(* IEC 61131-3 sources: 2026_Projet_YGO_ExcavatriceDragage/TOOLS/TEST_AUTO_CI/RESULTS/H_TREUILS_BENNE/reports (part 5) *)

    machine(HeartbeatIhmOk := TRUE, CanBusOperational := TRUE, JoyOperational := TRUE, CmdMode := E_Mode.DISABLE, TglJoystickMaster := TRUE, JoyRawY := 8000, CmdWinchSelect := 1);
    ADVANCE_TIME(20000000);
    machine(HeartbeatIhmOk := TRUE, CanBusOperational := TRUE, JoyOperational := TRUE, TglJoystickMaster := TRUE, JoyRawY := 8000, CmdWinchSelect := 1);
    ASSERT_TRUE(machine.BusOutputs.M1RelayFwd = FALSE, 'HARN-71: Enable=FALSE -> sorties sures');
    ASSERT_EQ(machine.M1_StepNumber, 0, 'HARN-71: palier neutralise');

    machine(HeartbeatIhmOk := TRUE, CanBusOperational := TRUE, JoyOperational := TRUE, CmdMode := E_Mode.MAINT_N1, TglJoystickMaster := TRUE, JoyRawY := 8000, CmdWinchSelect := 1);
    ADVANCE_TIME(50000000);
    machine(HeartbeatIhmOk := TRUE, CanBusOperational := TRUE, JoyOperational := TRUE, TglJoystickMaster := TRUE, JoyRawY := 8000, CmdWinchSelect := 1);
    (* ORACLE (main) : la reprise exige une NOUVELLE intention — l'adoption immédiate
       au ré-Enable = défaut D18 (rouge baseline attendu, cible T181-05) *)
    ASSERT_TRUE(machine.BusOutputs.M1RelayFwd = FALSE, 'HARN-71: pas de redemarrage auto au re-Enable (cible D18)');
END_TEST

TEST 'HARN-72 : Watchdog frein (retour frein ne suit pas) -> barriere coupe apres timeout'
    seqReqM1.RunRequest := FALSE; seqReqM1.ReqAscent := FALSE; seqReqM1.StepTgt := 0;
    seqReqM2.RunRequest := FALSE; seqReqM2.ReqAscent := FALSE; seqReqM2.StepTgt := 0;
    seqReqBucket.ExtractionControlActive := FALSE; seqReqBucket.DescendPermitDiveBucketOpen := FALSE;
    machine(HeartbeatIhmOk := TRUE, CanBusOperational := TRUE, JoyOperational := TRUE,
        CmdMode := E_Mode.MAINT_N1, CmdWinchSelect := 1, TglJoystickMaster := TRUE,
        SpeedTable := speedTable, ModelStepSpeedMps := modelSpeeds,
        SeqReqWinchM1 := seqReqM1, SeqReqWinchM2 := seqReqM2, SeqReqBucket := seqReqBucket,
        ModelSeedPosM1 := 2.0, ModelSeedPosM2 := 2.0, ModelReloadPositions := TRUE,
        ModelM2SpeedFactor := 1.0,
        ModelBrakeFeedbackFaultM1 := TRUE, (* retour frein M1 ne s ouvre jamais *)
        JoyRawX := 5000, JoyRawY := 5000, JoyDeadmanBtn := FALSE,
        EmergencyChainClosed := TRUE, PowerContactorEngaged := TRUE, HeartbeatIhmOk := TRUE
    );
    (* T181-00b : retour neutre sans commande >= 1500 ms pour purger RestartRequired/DeadTime *)
    machine(HeartbeatIhmOk := TRUE, CanBusOperational := TRUE, JoyOperational := TRUE, JoyDeadmanBtn := TRUE, TglJoystickMaster := TRUE, JoyRawY := 5000, CmdWinchSelect := 1, CmdMode := E_Mode.MAINT_N1);
    ADVANCE_TIME(2000000000);
    machine(HeartbeatIhmOk := TRUE, CanBusOperational := TRUE, JoyOperational := TRUE, JoyDeadmanBtn := TRUE, TglJoystickMaster := TRUE, JoyRawY := 5000, CmdWinchSelect := 1, CmdMode := E_Mode.MAINT_N1);
    machine(HeartbeatIhmOk := TRUE, CanBusOperational := TRUE, JoyOperational := TRUE, JoyDeadmanBtn := TRUE, TglJoystickMaster := TRUE, JoyRawY := 8000, CmdWinchSelect := 1, CmdMode := E_Mode.MAINT_N1);
    ADVANCE_TIME(5000000000); (* 5 s : tout timeout frein realiste a expire *)
    machine(HeartbeatIhmOk := TRUE, CanBusOperational := TRUE, JoyOperational := TRUE, TglJoystickMaster := TRUE, JoyRawY := 8000, CmdWinchSelect := 1, CmdMode := E_Mode.MAINT_N1);

    (* ORACLE (main) : frein incohérent -> la barrière coupe la commande de sens (TC-P10-012) *)
    ASSERT_TRUE(machine.BusWinch.WinchM1FinalInterlockRequest.RequestedRelayFwd, 'HARN-72: FB_Winch demande toujours le sens (defaut cote barriere)');
    ASSERT_TRUE(machine.BusOutputs.M1RelayFwd = FALSE, 'HARN-72: barriere a coupe (watchdog frein)');
    ASSERT_TRUE(machine.FinalInterlockGovernedM1, 'HARN-72: FinalInterlockGoverned TRUE');
END_TEST

TEST 'HARN-73 : Temps mort directionnel apres arret (inversion 200 ms) -> RelayRev retenu (CIBLE T175/T181-05)'
    seqReqM1.RunRequest := FALSE; seqReqM1.ReqAscent := FALSE; seqReqM1.StepTgt := 0;
    seqReqM2.RunRequest := FALSE; seqReqM2.ReqAscent := FALSE; seqReqM2.StepTgt := 0;
    seqReqBucket.ExtractionControlActive := FALSE; seqReqBucket.DescendPermitDiveBucketOpen := FALSE;
    machine(HeartbeatIhmOk := TRUE, CanBusOperational := TRUE, JoyOperational := TRUE,
        CmdMode := E_Mode.MAINT_N1, CmdWinchSelect := 1, TglJoystickMaster := TRUE,
        SpeedTable := speedTable, ModelStepSpeedMps := modelSpeeds,
        SeqReqWinchM1 := seqReqM1, SeqReqWinchM2 := seqReqM2, SeqReqBucket := seqReqBucket,
        ModelSeedPosM1 := 2.0, ModelSeedPosM2 := 2.0, ModelReloadPositions := TRUE,
        ModelM2SpeedFactor := 1.0,
        JoyRawX := 5000, JoyRawY := 5000, JoyDeadmanBtn := FALSE,
        EmergencyChainClosed := TRUE, PowerContactorEngaged := TRUE, HeartbeatIhmOk := TRUE
    );
    (* T181-00b : retour neutre sans commande >= 1500 ms pour purger RestartRequired/DeadTime *)
    machine(HeartbeatIhmOk := TRUE, CanBusOperational := TRUE, JoyOperational := TRUE, JoyDeadmanBtn := TRUE, TglJoystickMaster := TRUE, JoyRawY := 5000, CmdWinchSelect := 1, CmdMode := E_Mode.MAINT_N1);
    ADVANCE_TIME(2000000000);
    machine(HeartbeatIhmOk := TRUE, CanBusOperational := TRUE, JoyOperational := TRUE, JoyDeadmanBtn := TRUE, TglJoystickMaster := TRUE, JoyRawY := 5000, CmdWinchSelect := 1, CmdMode := E_Mode.MAINT_N1);
    machine(HeartbeatIhmOk := TRUE, CanBusOperational := TRUE, JoyOperational := TRUE, JoyDeadmanBtn := TRUE, TglJoystickMaster := TRUE, JoyRawY := 8000, CmdWinchSelect := 1, CmdMode := E_Mode.MAINT_N1);
    ADVANCE_TIME(200000000);
    machine(HeartbeatIhmOk := TRUE, CanBusOperational := TRUE, JoyOperational := TRUE, TglJoystickMaster := TRUE, JoyRawY := 8000, CmdWinchSelect := 1, CmdMode := E_Mode.MAINT_N1);
    machine(HeartbeatIhmOk := TRUE, CanBusOperational := TRUE, JoyOperational := TRUE, JoyDeadmanBtn := TRUE, TglJoystickMaster := TRUE, JoyRawY := 5000, CmdWinchSelect := 1, CmdMode := E_Mode.MAINT_N1);
    ADVANCE_TIME(20000000);
    machine(HeartbeatIhmOk := TRUE, CanBusOperational := TRUE, JoyOperational := TRUE, TglJoystickMaster := TRUE, JoyRawY := 5000, CmdWinchSelect := 1, CmdMode := E_Mode.MAINT_N1);
    (* Inversion 200 ms après l'arrêt *)
    machine(HeartbeatIhmOk := TRUE, CanBusOperational := TRUE, JoyOperational := TRUE, JoyDeadmanBtn := TRUE, TglJoystickMaster := TRUE, JoyRawY := 2000, CmdWinchSelect := 1, CmdMode := E_Mode.MAINT_N1);
    ADVANCE_TIME(200000000);
    machine(HeartbeatIhmOk := TRUE, CanBusOperational := TRUE, JoyOperational := TRUE, TglJoystickMaster := TRUE, JoyRawY := 2000, CmdWinchSelect := 1, CmdMode := E_Mode.MAINT_N1);

    (* PRECOND (durcissement T181-00b) : la barriere ne doit etre testee que si la demande de
       descente est REELlement presente en amont (RequestedRelayRev). Sans elle, M1RelayRev=FALSE
       est une tautologie (aucune demande a retenir). *)
    ASSERT_TRUE(machine.BusWinch.WinchM1FinalInterlockRequest.RequestedRelayRev, 'HARN-73: precondition - inversion descente reellement demandee');
    (* ORACLE (main) : délai interlock descente (400 ms) non écoulé -> la barriere retient RelayRev *)
    ASSERT_TRUE(machine.BusOutputs.M1RelayRev = FALSE, 'HARN-73: temps mort directionnel respecte (cible T175)');
END_TEST

TEST 'HARN-74a : Coast-down apres relache lourd -> PAS de faux PowerCutOff pendant la fenetre contacteurs (T178)'
    seqReqM1.RunRequest := FALSE; seqReqM1.ReqAscent := FALSE; seqReqM1.StepTgt := 0;
    seqReqM2.RunRequest := FALSE; seqReqM2.ReqAscent := FALSE; seqReqM2.StepTgt := 0;
    seqReqBucket.ExtractionControlActive := FALSE; seqReqBucket.DescendPermitDiveBucketOpen := FALSE;
    machine(HeartbeatIhmOk := TRUE, CanBusOperational := TRUE, JoyOperational := TRUE,
        CmdMode := E_Mode.MAINT_N1, CmdWinchSelect := 1, TglJoystickMaster := TRUE,
        SpeedTable := speedTable, ModelStepSpeedMps := modelSpeeds,
        SeqReqWinchM1 := seqReqM1, SeqReqWinchM2 := seqReqM2, SeqReqBucket := seqReqBucket,
        ModelSeedPosM1 := 2.0, ModelSeedPosM2 := 2.0, ModelReloadPositions := TRUE,
        ModelM2SpeedFactor := 1.0,
        JoyRawX := 5000, JoyRawY := 8000, JoyDeadmanBtn := FALSE,
        EmergencyChainClosed := TRUE, PowerContactorEngaged := TRUE, HeartbeatIhmOk := TRUE
    );
    (* T181-00b : retour neutre sans commande >= 1500 ms pour purger RestartRequired/DeadTime *)
    machine(HeartbeatIhmOk := TRUE, CanBusOperational := TRUE, JoyOperational := TRUE, JoyDeadmanBtn := TRUE, TglJoystickMaster := TRUE, JoyRawY := 5000, CmdWinchSelect := 1, CmdMode := E_Mode.MAINT_N1);
    ADVANCE_TIME(2000000000);
    machine(HeartbeatIhmOk := TRUE, CanBusOperational := TRUE, JoyOperational := TRUE, JoyDeadmanBtn := TRUE, TglJoystickMaster := TRUE, JoyRawY := 5000, CmdWinchSelect := 1, CmdMode := E_Mode.MAINT_N1);
    machine(HeartbeatIhmOk := TRUE, CanBusOperational := TRUE, JoyOperational := TRUE, JoyDeadmanBtn := TRUE, TglJoystickMaster := TRUE, JoyRawY := 8000, CmdWinchSelect := 1, CmdMode := E_Mode.MAINT_N1);
    ADVANCE_TIME(200000000);
    machine(HeartbeatIhmOk := TRUE, CanBusOperational := TRUE, JoyOperational := TRUE, TglJoystickMaster := TRUE, JoyRawY := 8000, CmdWinchSelect := 1, CmdMode := E_Mode.MAINT_N1);
    ASSERT_TRUE(machine.BusOutputs.M1RelayFwd, 'HARN-74a: precondition - montee plein pot');

    (* Relâche homme-mort plein déflexion : coast 500 ms (contacteurs pas encore retombés, v > 0) *)
    machine(HeartbeatIhmOk := TRUE, CanBusOperational := TRUE, JoyOperational := TRUE, JoyDeadmanBtn := FALSE, TglJoystickMaster := TRUE, JoyRawY := 8000, CmdWinchSelect := 1, CmdMode := E_Mode.MAINT_N1);
    ADVANCE_TIME(100000000); (* 100 ms au coeur de la fenêtre coast *)
    machine(HeartbeatIhmOk := TRUE, CanBusOperational := TRUE, JoyOperational := TRUE, TglJoystickMaster := TRUE, JoyRawY := 8000, CmdWinchSelect := 1, CmdMode := E_Mode.MAINT_N1);

    (* ORACLE (main) : pendant le coast — mouvement résiduel SANS commande : Méca A ne doit PAS armer *)
    ASSERT_TRUE(machine.BusWinch.WinchM1Safety.PowerCutOff = FALSE, 'HARN-74a: PAS de faux PowerCutOff pendant le coast (T178)');
    ASSERT_TRUE(machine.BusWinch.WinchM1Safety.SafeStop = FALSE, 'HARN-74a: PAS de SafeStop pendant le coast (Meca A)');
END_TEST

TEST 'HARN-74b : Coast-down prolonge -> Meca B arme a 3 s (CIBLE T178, ROUGE baseline)'
    seqReqM1.RunRequest := FALSE; seqReqM1.ReqAscent := FALSE; seqReqM1.StepTgt := 0;
    seqReqM2.RunRequest := FALSE; seqReqM2.ReqAscent := FALSE; seqReqM2.StepTgt := 0;
    seqReqBucket.ExtractionControlActive := FALSE; seqReqBucket.DescendPermitDiveBucketOpen := FALSE;
    machine(HeartbeatIhmOk := TRUE, CanBusOperational := TRUE, JoyOperational := TRUE,
        CmdMode := E_Mode.MAINT_N1, CmdWinchSelect := 1, TglJoystickMaster := TRUE,
        SpeedTable := speedTable, ModelStepSpeedMps := modelSpeeds,
        SeqReqWinchM1 := seqReqM1, SeqReqWinchM2 := seqReqM2, SeqReqBucket := seqReqBucket,
        ModelSeedPosM1 := 2.0, ModelSeedPosM2 := 2.0, ModelReloadPositions := TRUE,
        ModelM2SpeedFactor := 1.0,
        JoyRawX := 5000, JoyRawY := 8000, JoyDeadmanBtn := FALSE,
        EmergencyChainClosed := TRUE, PowerContactorEngaged := TRUE, HeartbeatIhmOk := TRUE
    );
    (* T181-00b : retour neutre sans commande >= 1500 ms pour purger RestartRequired/DeadTime *)
    machine(HeartbeatIhmOk := TRUE, CanBusOperational := TRUE, JoyOperational := TRUE, JoyDeadmanBtn := TRUE, TglJoystickMaster := TRUE, JoyRawY := 5000, CmdWinchSelect := 1, CmdMode := E_Mode.MAINT_N1);
    ADVANCE_TIME(2000000000);
    machine(HeartbeatIhmOk := TRUE, CanBusOperational := TRUE, JoyOperational := TRUE, JoyDeadmanBtn := TRUE, TglJoystickMaster := TRUE, JoyRawY := 5000, CmdWinchSelect := 1, CmdMode := E_Mode.MAINT_N1);
    machine(HeartbeatIhmOk := TRUE, CanBusOperational := TRUE, JoyOperational := TRUE, JoyDeadmanBtn := TRUE, TglJoystickMaster := TRUE, JoyRawY := 8000, CmdWinchSelect := 1, CmdMode := E_Mode.MAINT_N1);
    ADVANCE_TIME(200000000);
    machine(HeartbeatIhmOk := TRUE, CanBusOperational := TRUE, JoyOperational := TRUE, TglJoystickMaster := TRUE, JoyRawY := 8000, CmdWinchSelect := 1, CmdMode := E_Mode.MAINT_N1);
    machine(HeartbeatIhmOk := TRUE, CanBusOperational := TRUE, JoyOperational := TRUE, JoyDeadmanBtn := FALSE, TglJoystickMaster := TRUE, JoyRawY := 8000, CmdWinchSelect := 1, CmdMode := E_Mode.MAINT_N1);
    ADVANCE_TIME(4000000000); (* 4 s > 3 s *)
    machine(HeartbeatIhmOk := TRUE, CanBusOperational := TRUE, JoyOperational := TRUE, TglJoystickMaster := TRUE, JoyRawY := 8000, CmdWinchSelect := 1, CmdMode := E_Mode.MAINT_N1);
    (* ORACLE (main) : Méca B (absence confirmation arrêt) arme à 3 s -> SafeStop *)
    ASSERT_TRUE(machine.BusWinch.WinchM1Safety.SafeStop, 'HARN-74b: Meca B arme a 3 s (cible T178)');
END_TEST

TEST 'HARN-75 : Redemarrage a chaud (FirstScanDone) -> temps mort directionnel NON bypassse (D18, ROUGE baseline)'
    (* Scénario D18 : direction ≠ 0 maintenue à travers une ré-init (Enable FALSE->TRUE) ;
       l'interlock directionnel doit s'appliquer au front montant Enable — PAS via FirstScanDone. *)
    seqReqM1.RunRequest := FALSE; seqReqM1.ReqAscent := FALSE; seqReqM1.StepTgt := 0;
    seqReqM2.RunRequest := FALSE; seqReqM2.ReqAscent := FALSE; seqReqM2.StepTgt := 0;
    seqReqBucket.ExtractionControlActive := FALSE; seqReqBucket.DescendPermitDiveBucketOpen := FALSE;
    machine(HeartbeatIhmOk := TRUE, CanBusOperational := TRUE, JoyOperational := TRUE,
        CmdMode := E_Mode.MAINT_N1, CmdWinchSelect := 1, TglJoystickMaster := TRUE,
        SpeedTable := speedTable, ModelStepSpeedMps := modelSpeeds,
        SeqReqWinchM1 := seqReqM1, SeqReqWinchM2 := seqReqM2, SeqReqBucket := seqReqBucket,
        ModelSeedPosM1 := 2.0, ModelSeedPosM2 := 2.0, ModelReloadPositions := TRUE,
        ModelM2SpeedFactor := 1.0,
        JoyRawX := 5000, JoyRawY := 8000, JoyDeadmanBtn := FALSE,
        EmergencyChainClosed := TRUE, PowerContactorEngaged := TRUE, HeartbeatIhmOk := TRUE
    );
    (* T181-00b : retour neutre sans commande >= 1500 ms pour purger RestartRequired/DeadTime *)
    machine(HeartbeatIhmOk := TRUE, CanBusOperational := TRUE, JoyOperational := TRUE, JoyDeadmanBtn := TRUE, TglJoystickMaster := TRUE, JoyRawY := 5000, CmdWinchSelect := 1, CmdMode := E_Mode.MAINT_N1);
    ADVANCE_TIME(2000000000);
    machine(HeartbeatIhmOk := TRUE, CanBusOperational := TRUE, JoyOperational := TRUE, JoyDeadmanBtn := TRUE, TglJoystickMaster := TRUE, JoyRawY := 5000, CmdWinchSelect := 1, CmdMode := E_Mode.MAINT_N1);
    machine(HeartbeatIhmOk := TRUE, CanBusOperational := TRUE, JoyOperational := TRUE, JoyDeadmanBtn := TRUE, TglJoystickMaster := TRUE, JoyRawY := 8000, CmdWinchSelect := 1, CmdMode := E_Mode.MAINT_N1);
    ADVANCE_TIME(200000000);
    machine(HeartbeatIhmOk := TRUE, CanBusOperational := TRUE, JoyOperational := TRUE, TglJoystickMaster := TRUE, JoyRawY := 8000, CmdWinchSelect := 1, CmdMode := E_Mode.MAINT_N1);
    ASSERT_TRUE(machine.BusOutputs.M1RelayFwd, 'HARN-75: precondition - montee active');

    machine(HeartbeatIhmOk := TRUE, CanBusOperational := TRUE, JoyOperational := TRUE, CmdMode := E_Mode.DISABLE, TglJoystickMaster := TRUE, JoyRawY := 8000, CmdWinchSelect := 1);
    ADVANCE_TIME(20000000);
    machine(HeartbeatIhmOk := TRUE, CanBusOperational := TRUE, JoyOperational := TRUE, CmdMode := E_Mode.MAINT_N1, TglJoystickMaster := TRUE, JoyRawY := 8000, CmdWinchSelect := 1);
    ADVANCE_TIME(100000000);
    machine(HeartbeatIhmOk := TRUE, CanBusOperational := TRUE, JoyOperational := TRUE, TglJoystickMaster := TRUE, JoyRawY := 8000, CmdWinchSelect := 1, CmdMode := E_Mode.MAINT_N1);

    (* ORACLE (main) : après hot-restart avec direction maintenue, un signal D18 REEL
       (DirectionChangePending ou FinalRestartInhibit) doit etre pose. Retire l'echappatoire
       "OR M1RelayFwd=FALSE" qui rendait l'assertion vraie par defaut (faux vert D18). *)
    ASSERT_TRUE(machine.BusWinch.WinchM1State.DirectionChangePending
                OR machine.BusWinch.WinchM1State.FinalRestartInhibit,
                'HARN-75: temps mort applique au hot-restart (D18, cible T181-05)');
END_TEST

(* ═══════════════ FAMILLE 8 — Croisement audit T180 (HARN-8x) ═══════════════ *)

TEST 'HARN-80 : CAS-001 retombee contacteur EN MARCHE (feedback incoherent) -> defaut + neutralisation (CIBLE T180)'
    seqReqM1.RunRequest := FALSE; seqReqM1.ReqAscent := FALSE; seqReqM1.StepTgt := 0;
    seqReqM2.RunRequest := FALSE; seqReqM2.ReqAscent := FALSE; seqReqM2.StepTgt := 0;
    seqReqBucket.ExtractionControlActive := FALSE; seqReqBucket.DescendPermitDiveBucketOpen := FALSE;
    machine(HeartbeatIhmOk := TRUE, CanBusOperational := TRUE, JoyOperational := TRUE,
        CmdMode := E_Mode.MAINT_N1, CmdWinchSelect := 1, TglJoystickMaster := TRUE,
        SpeedTable := speedTable, ModelStepSpeedMps := modelSpeeds,
        SeqReqWinchM1 := seqReqM1, SeqReqWinchM2 := seqReqM2, SeqReqBucket := seqReqBucket,
        ModelSeedPosM1 := 2.0, ModelSeedPosM2 := 2.0, ModelReloadPositions := TRUE,
        ModelM2SpeedFactor := 1.0,
        ModelContactorsReleaseFaultM1 := TRUE, (* contacteurs declares retombes ALORS qu on commande *)
        JoyRawX := 5000, JoyRawY := 8000, JoyDeadmanBtn := FALSE,
        EmergencyChainClosed := TRUE, PowerContactorEngaged := TRUE, HeartbeatIhmOk := TRUE
    );
    (* T181-00b : retour neutre sans commande >= 1500 ms pour purger RestartRequired/DeadTime *)
    machine(HeartbeatIhmOk := TRUE, CanBusOperational := TRUE, JoyOperational := TRUE, JoyDeadmanBtn := TRUE, TglJoystickMaster := TRUE, JoyRawY := 5000, CmdWinchSelect := 1, CmdMode := E_Mode.MAINT_N1);
    ADVANCE_TIME(2000000000);
    machine(HeartbeatIhmOk := TRUE, CanBusOperational := TRUE, JoyOperational := TRUE, JoyDeadmanBtn := TRUE, TglJoystickMaster := TRUE, JoyRawY := 5000, CmdWinchSelect := 1, CmdMode := E_Mode.MAINT_N1);
    machine(HeartbeatIhmOk := TRUE, CanBusOperational := TRUE, JoyOperational := TRUE, JoyDeadmanBtn := TRUE, TglJoystickMaster := TRUE, JoyRawY := 8000, CmdWinchSelect := 1, CmdMode := E_Mode.MAINT_N1);
    ADVANCE_TIME(300000000);
    machine(HeartbeatIhmOk := TRUE, CanBusOperational := TRUE, JoyOperational := TRUE, TglJoystickMaster := TRUE, JoyRawY := 8000, CmdWinchSelect := 1, CmdMode := E_Mode.MAINT_N1);

    (* PRECOND (durcissement T181-00b) : le defaut CAS-001 ne se teste qu en montee REELlement
       commandee (sinon RelayFwd=FALSE est une tautologie : rien ne bouge -> rien a neutraliser). *)
    ASSERT_TRUE(machine.BusOutputs.M1RelayFwd, 'HARN-80: precondition - montee M1 commandee');
    (* ORACLE (main) : en marche, retombee contacteur incoherente -> defaut Error DETECTE.
       Retire "OR RelayFwd=FALSE" (vrai par defaut). CAS-001 / T180. *)
    ASSERT_TRUE(machine.BusWinch.WinchM1Safety.Error, 'HARN-80: CAS-001 detecte (defaut Error, cible T180)');
END_TEST

TEST 'HARN-81 : CAS-012 demande benne pendant mouvement treuil -> demande REFUSEE (CIBLE T175 AC3)'
    seqReqM1.RunRequest := FALSE; seqReqM1.ReqAscent := FALSE; seqReqM1.StepTgt := 0;
    seqReqM2.RunRequest := FALSE; seqReqM2.ReqAscent := FALSE; seqReqM2.StepTgt := 0;
    seqReqBucket.ExtractionControlActive := FALSE; seqReqBucket.DescendPermitDiveBucketOpen := FALSE;
    machine(HeartbeatIhmOk := TRUE, CanBusOperational := TRUE, JoyOperational := TRUE,
        CmdMode := E_Mode.MAINT_N1, CmdWinchSelect := 0, TglJoystickMaster := TRUE,
        SpeedTable := speedTable, ModelStepSpeedMps := modelSpeeds,
        SeqReqWinchM1 := seqReqM1, SeqReqWinchM2 := seqReqM2, SeqReqBucket := seqReqBucket,
        ModelSeedPosM1 := 2.0, ModelSeedPosM2 := 2.0, ModelReloadPositions := TRUE,
        ModelM2SpeedFactor := 1.0,
        JoyRawX := 5000, JoyRawY := 5000, JoyDeadmanBtn := FALSE,
        BucketCmdOpen := FALSE, BucketCmdClose := FALSE,
        EmergencyChainClosed := TRUE, PowerContactorEngaged := TRUE, HeartbeatIhmOk := TRUE
    );
    machine(HeartbeatIhmOk := TRUE, CanBusOperational := TRUE, JoyOperational := TRUE, JoyDeadmanBtn := TRUE, TglJoystickMaster := TRUE, CmdWinchSelect := 0, CmdMode := E_Mode.MAINT_N1);
    (* T181-00b : retour neutre sans commande >= 1500 ms pour purger RestartRequired/DeadTime *)
    ADVANCE_TIME(2000000000);
    machine(HeartbeatIhmOk := TRUE, CanBusOperational := TRUE, JoyOperational := TRUE, JoyDeadmanBtn := TRUE, TglJoystickMaster := TRUE, CmdWinchSelect := 0, CmdMode := E_Mode.MAINT_N1);
    machine(HeartbeatIhmOk := TRUE, CanBusOperational := TRUE, JoyOperational := TRUE, JoyDeadmanBtn := TRUE, TglJoystickMaster := TRUE, JoyRawY := 8000, CmdWinchSelect := 0, CmdMode := E_Mode.MAINT_N1);
    ADVANCE_TIME(200000000);
    machine(HeartbeatIhmOk := TRUE, CanBusOperational := TRUE, JoyOperational := TRUE, TglJoystickMaster := TRUE, JoyRawY := 8000, CmdWinchSelect := 0, CmdMode := E_Mode.MAINT_N1);
    ASSERT_TRUE(machine.M1_StepNumber > 0, 'HARN-81: precondition - treuils en mouvement');

    machine(HeartbeatIhmOk := TRUE, CanBusOperational := TRUE, JoyOperational := TRUE, BucketCmdClose := TRUE, JoyDeadmanBtn := TRUE, TglJoystickMaster := TRUE, JoyRawY := 8000, CmdWinchSelect := 0, CmdMode := E_Mode.MAINT_N1);
    ADVANCE_TIME(50000000);
    machine(HeartbeatIhmOk := TRUE, CanBusOperational := TRUE, JoyOperational := TRUE, BucketCmdClose := TRUE, TglJoystickMaster := TRUE, JoyRawY := 8000, CmdWinchSelect := 0, CmdMode := E_Mode.MAINT_N1);

    (* ORACLE (main) : anti-traversée — la demande benne est refusée tant que les treuils agissent *)
    ASSERT_TRUE(machine.BusWinch.BucketBusy = FALSE, 'HARN-81: CAS-012 demande benne refusee (cible T175 AC3)');
END_TEST

TEST 'HARN-82 : CAS-002 AU pendant transition d etape -> coupure propre, pas d etat incoherent au rearmement'
    seqReqM1.RunRequest := FALSE; seqReqM1.ReqAscent := FALSE; seqReqM1.StepTgt := 0;
    seqReqM2.RunRequest := FALSE; seqReqM2.ReqAscent := FALSE; seqReqM2.StepTgt := 0;
    seqReqBucket.ExtractionControlActive := FALSE; seqReqBucket.DescendPermitDiveBucketOpen := FALSE;
    machine(HeartbeatIhmOk := TRUE, CanBusOperational := TRUE, JoyOperational := TRUE,
        CmdMode := E_Mode.SEMI_AUTO, CmdWinchSelect := 0,
        SpeedTable := speedTable, ModelStepSpeedMps := modelSpeeds,
        SeqReqWinchM1 := seqReqM1, SeqReqWinchM2 := seqReqM2, SeqReqBucket := seqReqBucket,
        ModelSeedPosM1 := 2.0, ModelSeedPosM2 := 2.0, ModelReloadPositions := TRUE,
        ModelM2SpeedFactor := 1.0,
        JoyRawX := 5000, JoyRawY := 5000, JoyDeadmanBtn := FALSE,
        EmergencyChainClosed := TRUE, PowerContactorEngaged := TRUE, HeartbeatIhmOk := TRUE
    );
    machine(HeartbeatIhmOk := TRUE, CanBusOperational := TRUE, JoyOperational := TRUE, ModelReloadPositions := FALSE, CmdMode := E_Mode.SEMI_AUTO);
    (* T181-00b : retour neutre sans commande >= 1500 ms pour purger RestartRequired/DeadTime *)
    machine(HeartbeatIhmOk := TRUE, CanBusOperational := TRUE, JoyOperational := TRUE, CmdMode := E_Mode.SEMI_AUTO, JoyDeadmanBtn := TRUE, EmergencyChainClosed := TRUE, PowerContactorEngaged := TRUE);
    ADVANCE_TIME(2000000000);
    machine(HeartbeatIhmOk := TRUE, CanBusOperational := TRUE, JoyOperational := TRUE, CmdMode := E_Mode.SEMI_AUTO, JoyDeadmanBtn := TRUE, EmergencyChainClosed := TRUE, PowerContactorEngaged := TRUE);
    seqReqM1.RunRequest := TRUE; seqReqM1.ReqAscent := TRUE; seqReqM1.ReqDescend := FALSE; seqReqM1.StepTgt := 3;
    seqReqM2.RunRequest := TRUE; seqReqM2.ReqAscent := TRUE; seqReqM2.ReqDescend := FALSE; seqReqM2.StepTgt := 3;
    machine(HeartbeatIhmOk := TRUE, CanBusOperational := TRUE, JoyOperational := TRUE, SeqReqWinchM1 := seqReqM1, SeqReqWinchM2 := seqReqM2, SeqReqBucket := seqReqBucket,
        CmdMode := E_Mode.SEMI_AUTO, JoyRawX := 5000, JoyRawY := 5000, JoyDeadmanBtn := TRUE,
        EmergencyChainClosed := TRUE, PowerContactorEngaged := TRUE, HeartbeatIhmOk := TRUE);
    ADVANCE_TIME(200000000);
    machine(HeartbeatIhmOk := TRUE, CanBusOperational := TRUE, JoyOperational := TRUE, SeqReqWinchM1 := seqReqM1, SeqReqWinchM2 := seqReqM2, SeqReqBucket := seqReqBucket,
        CmdMode := E_Mode.SEMI_AUTO, JoyRawX := 5000, JoyRawY := 5000, JoyDeadmanBtn := TRUE,
        EmergencyChainClosed := TRUE, PowerContactorEngaged := TRUE, HeartbeatIhmOk := TRUE);
    ASSERT_TRUE(machine.BusOutputs.M1RelayFwd, 'HARN-82: precondition - mouvement semi-auto');

    machine(HeartbeatIhmOk := TRUE, CanBusOperational := TRUE, JoyOperational := TRUE, EmergencyChainClosed := FALSE, PowerContactorEngaged := FALSE);
    ADVANCE_TIME(50000000);
    machine(HeartbeatIhmOk := TRUE, CanBusOperational := TRUE, JoyOperational := TRUE, SeqReqWinchM1 := seqReqM1, SeqReqWinchM2 := seqReqM2, SeqReqBucket := seqReqBucket,
        CmdMode := E_Mode.SEMI_AUTO, JoyRawX := 5000, JoyRawY := 5000, JoyDeadmanBtn := TRUE,
        EmergencyChainClosed := TRUE, PowerContactorEngaged := TRUE, HeartbeatIhmOk := TRUE);
    ASSERT_TRUE(machine.BusOutputs.M1RelayFwd = FALSE, 'HARN-82: coupure propre a l AU');

    seqReqM1.RunRequest := FALSE; seqReqM2.RunRequest := FALSE;
    machine(CanBusOperational := TRUE, JoyOperational := TRUE, EmergencyChainClosed := TRUE, PowerContactorEngaged := TRUE, HeartbeatIhmOk := TRUE, BtnResetMachine := TRUE,
            SeqReqWinchM1 := seqReqM1, SeqReqWinchM2 := seqReqM2, SeqReqBucket := seqReqBucket);
    ADVANCE_TIME(10000000);
    machine(HeartbeatIhmOk := TRUE, CanBusOperational := TRUE, JoyOperational := TRUE, BtnResetMachine := FALSE, SeqReqWinchM1 := seqReqM1, SeqReqWinchM2 := seqReqM2, SeqReqBucket := seqReqBucket);
    ADVANCE_TIME(100000000);
    machine(HeartbeatIhmOk := TRUE, CanBusOperational := TRUE, JoyOperational := TRUE, SeqReqWinchM1 := seqReqM1, SeqReqWinchM2 := seqReqM2, SeqReqBucket := seqReqBucket,
        CmdMode := E_Mode.SEMI_AUTO, JoyRawX := 5000, JoyRawY := 5000, JoyDeadmanBtn := TRUE,
        EmergencyChainClosed := TRUE, PowerContactorEngaged := TRUE, HeartbeatIhmOk := TRUE);

    (* ORACLE (main) : après réarmement, aucune reprise sans ordre explicite *)
    ASSERT_TRUE(machine.BusOutputs.M1RelayFwd = FALSE, 'HARN-82: pas de reprise apres rearmement sans ordre');
    ASSERT_TRUE(machine.BusOutputs.M2RelayFwd = FALSE, 'HARN-82: idem M2');
    ASSERT_EQ(machine.M1_StepNumber, 0, 'HARN-82: etat coherent (palier 0)');
END_TEST
